(* IEC 61131-3 sources: virtual-bottling-plant/plc/src/generated/io, 9 files *)

(* ---- IO_C501.st ---- *)
(* GENERATED by plc/scripts/gen_plc_io.py from contracts/modbus/sim-io.yaml. Do not edit by hand. *)
(* Remote I/O station C501 (Modbus unit 5). *)
PROGRAM IO_C501
  VAR_EXTERNAL
    G_In : ST_SimInputs;
    G_Out : ST_SimOutputs;
  END_VAR
  VAR
    C501_Running AT %IX100.7 : BOOL;
    C501_Jam AT %IX101.0 : BOOL;
    C501_Breakdown AT %IX101.1 : BOOL;
    LSL502_CapsEmpty AT %IX101.2 : BOOL;
    C501_Run AT %QX101.2 : BOOL;
    C501_Speed AT %IW120 : UINT;
    C501_Count_HI AT %IW121 : UINT;
    C501_Count_LO AT %IW122 : UINT;
    C501_Torque AT %IW123 : UINT;
    LT502_CapHopper AT %IW124 : UINT;
    C501_Heartbeat AT %IW125 : UINT;
    C501_SpeedSP AT %QW104 : UINT;
  END_VAR
  G_In.C501_Running := C501_Running;
  G_In.C501_Jam := C501_Jam;
  G_In.C501_Breakdown := C501_Breakdown;
  G_In.LSL502_CapsEmpty := LSL502_CapsEmpty;
  C501_Run := G_Out.C501_Run;
  G_In.C501_Speed := UINT_TO_REAL(C501_Speed);
  G_In.C501_Count := UINT_TO_UDINT(C501_Count_HI) * 65536 + UINT_TO_UDINT(C501_Count_LO);
  G_In.C501_Torque := UINT_TO_REAL(C501_Torque) / 100.0;
  G_In.LT502_CapHopper := UINT_TO_REAL(LT502_CapHopper) / 10.0;
  G_In.C501_Heartbeat := C501_Heartbeat;
  C501_SpeedSP := REAL_TO_UINT(LIMIT(0.0, G_Out.C501_SpeedSP, 65535.0));
END_PROGRAM

(* ---- IO_F401.st ---- *)
(* GENERATED by plc/scripts/gen_plc_io.py from contracts/modbus/sim-io.yaml. Do not edit by hand. *)
(* Remote I/O station F401 (Modbus unit 4). *)
PROGRAM IO_F401
  VAR_EXTERNAL
    G_In : ST_SimInputs;
    G_Out : ST_SimOutputs;
  END_VAR
  VAR
    F401_Running AT %IX100.5 : BOOL;
    F401_NozzleLeak AT %IX100.6 : BOOL;
    F401_Run AT %QX101.1 : BOOL;
    F401_Speed AT %IW116 : UINT;
    F401_Count_HI AT %IW117 : UINT;
    F401_Count_LO AT %IW118 : UINT;
    F401_Heartbeat AT %IW119 : UINT;
    F401_SpeedSP AT %QW102 : UINT;
    F401_FillTargetG AT %QW103 : UINT;
  END_VAR
  G_In.F401_Running := F401_Running;
  G_In.F401_NozzleLeak := F401_NozzleLeak;
  F401_Run := G_Out.F401_Run;
  G_In.F401_Speed := UINT_TO_REAL(F401_Speed);
  G_In.F401_Count := UINT_TO_UDINT(F401_Count_HI) * 65536 + UINT_TO_UDINT(F401_Count_LO);
  G_In.F401_Heartbeat := F401_Heartbeat;
  F401_SpeedSP := REAL_TO_UINT(LIMIT(0.0, G_Out.F401_SpeedSP, 65535.0));
  F401_FillTargetG := REAL_TO_UINT(LIMIT(0.0, G_Out.F401_FillTargetG * 10.0, 65535.0));
END_PROGRAM

(* ---- IO_K801.st ---- *)
(* GENERATED by plc/scripts/gen_plc_io.py from contracts/modbus/sim-io.yaml. Do not edit by hand. *)
(* Remote I/O station K801 (Modbus unit 8). *)
PROGRAM IO_K801
  VAR_EXTERNAL
    G_In : ST_SimInputs;
    G_Out : ST_SimOutputs;
  END_VAR
  VAR
    K801_Running AT %IX102.0 : BOOL;
    K801_Jam AT %IX102.1 : BOOL;
    K801_Breakdown AT %IX102.2 : BOOL;
    K801_Run AT %QX101.5 : BOOL;
    K801_Speed AT %IW177 : UINT;
    K801_CaseCount_HI AT %IW178 : UINT;
    K801_CaseCount_LO AT %IW179 : UINT;
    K801_Heartbeat AT %IW180 : UINT;
    K801_SpeedSP AT %QW108 : UINT;
  END_VAR
  G_In.K801_Running := K801_Running;
  G_In.K801_Jam := K801_Jam;
  G_In.K801_Breakdown := K801_Breakdown;
  K801_Run := G_Out.K801_Run;
  G_In.K801_Speed := UINT_TO_REAL(K801_Speed);
  G_In.K801_CaseCount := UINT_TO_UDINT(K801_CaseCount_HI) * 65536 + UINT_TO_UDINT(K801_CaseCount_LO);
  G_In.K801_Heartbeat := K801_Heartbeat;
  K801_SpeedSP := REAL_TO_UINT(LIMIT(0.0, G_Out.K801_SpeedSP, 65535.0));
END_PROGRAM

(* ---- IO_L601.st ---- *)
(* GENERATED by plc/scripts/gen_plc_io.py from contracts/modbus/sim-io.yaml. Do not edit by hand. *)
(* Remote I/O station L601 (Modbus unit 6). *)
PROGRAM IO_L601
  VAR_EXTERNAL
    G_In : ST_SimInputs;
    G_Out : ST_SimOutputs;
  END_VAR
  VAR
    L601_Running AT %IX101.3 : BOOL;
    L601_RollEmpty AT %IX101.4 : BOOL;
    L601_LabelError AT %IX101.5 : BOOL;
    L601_Breakdown AT %IX101.6 : BOOL;
    L601_Run AT %QX101.3 : BOOL;
    L601_Speed AT %IW126 : UINT;
    L601_Count_HI AT %IW127 : UINT;
    L601_Count_LO AT %IW128 : UINT;
    L601_RollRemaining AT %IW129 : UINT;
    L601_Heartbeat AT %IW130 : UINT;
    L601_SpeedSP AT %QW105 : UINT;
  END_VAR
  G_In.L601_Running := L601_Running;
  G_In.L601_RollEmpty := L601_RollEmpty;
  G_In.L601_LabelError := L601_LabelError;
  G_In.L601_Breakdown := L601_Breakdown;
  L601_Run := G_Out.L601_Run;
  G_In.L601_Speed := UINT_TO_REAL(L601_Speed);
  G_In.L601_Count := UINT_TO_UDINT(L601_Count_HI) * 65536 + UINT_TO_UDINT(L601_Count_LO);
  G_In.L601_RollRemaining := UINT_TO_REAL(L601_RollRemaining);
  G_In.L601_Heartbeat := L601_Heartbeat;
  L601_SpeedSP := REAL_TO_UINT(LIMIT(0.0, G_Out.L601_SpeedSP, 65535.0));
END_PROGRAM

(* ---- IO_LINE.st ---- *)
(* GENERATED by plc/scripts/gen_plc_io.py from contracts/modbus/sim-io.yaml. Do not edit by hand. *)
(* Remote I/O station LINE (Modbus unit 9). *)
PROGRAM IO_LINE
  VAR_EXTERNAL
    G_In : ST_SimInputs;
  END_VAR
  VAR
    CV1_Full AT %IX102.3 : BOOL;
    CV2_Full AT %IX102.4 : BOOL;
    CV3_Full AT %IX102.5 : BOOL;
    CV4_Full AT %IX102.6 : BOOL;
    PB_Start AT %IX102.7 : BOOL;
    PB_Stop AT %IX103.0 : BOOL;
    PB_Reset AT %IX103.1 : BOOL;
    SIM_TimeMs_HI AT %IW181 : UINT;
    SIM_TimeMs_LO AT %IW182 : UINT;
    CV1_Fill AT %IW183 : UINT;
    CV2_Fill AT %IW184 : UINT;
    CV3_Fill AT %IW185 : UINT;
    CV4_Fill AT %IW186 : UINT;
    LINE_Heartbeat AT %IW187 : UINT;
  END_VAR
  G_In.CV1_Full := CV1_Full;
  G_In.CV2_Full := CV2_Full;
  G_In.CV3_Full := CV3_Full;
  G_In.CV4_Full := CV4_Full;
  G_In.PB_Start := PB_Start;
  G_In.PB_Stop := PB_Stop;
  G_In.PB_Reset := PB_Reset;
  G_In.SIM_TimeMs := UINT_TO_UDINT(SIM_TimeMs_HI) * 65536 + UINT_TO_UDINT(SIM_TimeMs_LO);
  G_In.CV1_Fill := UINT_TO_REAL(CV1_Fill);
  G_In.CV2_Fill := UINT_TO_REAL(CV2_Fill);
  G_In.CV3_Fill := UINT_TO_REAL(CV3_Fill);
  G_In.CV4_Fill := UINT_TO_REAL(CV4_Fill);
  G_In.LINE_Heartbeat := LINE_Heartbeat;
END_PROGRAM

(* ---- IO_P201.st ---- *)
(* GENERATED by plc/scripts/gen_plc_io.py from contracts/modbus/sim-io.yaml. Do not edit by hand. *)
(* Remote I/O station P201 (Modbus unit 2). *)
PROGRAM IO_P201
  VAR_EXTERNAL
    G_In : ST_SimInputs;
    G_Out : ST_SimOutputs;
  END_VAR
  VAR
    ZS203_DivertOpen AT %IX100.3 : BOOL;
    XV203_Divert AT %QX100.7 : BOOL;
    TT201_InTemp AT %IW109 : UINT;
    TT202_OutTemp AT %IW110 : UINT;
    FT201_Flow AT %IW111 : UINT;
    PT201_SteamPressure AT %IW112 : UINT;
    P201_Heartbeat AT %IW113 : UINT;
    TCV201_SteamValve AT %QW101 : UINT;
  END_VAR
  G_In.ZS203_DivertOpen := ZS203_DivertOpen;
  XV203_Divert := G_Out.XV203_Divert;
  G_In.TT201_InTemp := UINT_TO_REAL(TT201_InTemp) / 10.0;
  G_In.TT202_OutTemp := UINT_TO_REAL(TT202_OutTemp) / 10.0;
  G_In.FT201_Flow := UINT_TO_REAL(FT201_Flow);
  G_In.PT201_SteamPressure := UINT_TO_REAL(PT201_SteamPressure) / 100.0;
  G_In.P201_Heartbeat := P201_Heartbeat;
  TCV201_SteamValve := REAL_TO_UINT(LIMIT(0.0, G_Out.TCV201_SteamValve * 10.0, 65535.0));
END_PROGRAM

(* ---- IO_Q701.st ---- *)
(* GENERATED by plc/scripts/gen_plc_io.py from contracts/modbus/sim-io.yaml. Do not edit by hand. *)
(* Remote I/O station Q701 (Modbus unit 7). *)
PROGRAM IO_Q701
  VAR_EXTERNAL
    G_In : ST_SimInputs;
    G_Out : ST_SimOutputs;
  END_VAR
  VAR
    Q701_Running AT %IX101.7 : BOOL;
    Q701_Run AT %QX101.4 : BOOL;
    Q701_Speed AT %IW131 : UINT;
    Q701_Count_HI AT %IW132 : UINT;
    Q701_Count_LO AT %IW133 : UINT;
    Q701_RejectCount_HI AT %IW134 : UINT;
    Q701_RejectCount_LO AT %IW135 : UINT;
    WT701_LastWeight AT %IW136 : UINT;
    Q701_Heartbeat AT %IW137 : UINT;
    Q701_N01_Seq AT %IW141 : UINT;
    Q701_N01_Mean AT %IW142 : UINT;
    Q701_N01_Range AT %IW143 : UINT;
    Q701_N02_Seq AT %IW144 : UINT;
    Q701_N02_Mean AT %IW145 : UINT;
    Q701_N02_Range AT %IW146 : UINT;
    Q701_N03_Seq AT %IW147 : UINT;
    Q701_N03_Mean AT %IW148 : UINT;
    Q701_N03_Range AT %IW149 : UINT;
    Q701_N04_Seq AT %IW150 : UINT;
    Q701_N04_Mean AT %IW151 : UINT;
    Q701_N04_Range AT %IW152 : UINT;
    Q701_N05_Seq AT %IW153 : UINT;
    Q701_N05_Mean AT %IW154 : UINT;
    Q701_N05_Range AT %IW155 : UINT;
    Q701_N06_Seq AT %IW156 : UINT;
    Q701_N06_Mean AT %IW157 : UINT;
    Q701_N06_Range AT %IW158 : UINT;
    Q701_N07_Seq AT %IW159 : UINT;
    Q701_N07_Mean AT %IW160 : UINT;
    Q701_N07_Range AT %IW161 : UINT;
    Q701_N08_Seq AT %IW162 : UINT;
    Q701_N08_Mean AT %IW163 : UINT;
    Q701_N08_Range AT %IW164 : UINT;
    Q701_N09_Seq AT %IW165 : UINT;
    Q701_N09_Mean AT %IW166 : UINT;
    Q701_N09_Range AT %IW167 : UINT;
    Q701_N10_Seq AT %IW168 : UINT;
    Q701_N10_Mean AT %IW169 : UINT;
    Q701_N10_Range AT %IW170 : UINT;
    Q701_N11_Seq AT %IW171 : UINT;
    Q701_N11_Mean AT %IW172 : UINT;
    Q701_N11_Range AT %IW173 : UINT;
    Q701_N12_Seq AT %IW174 : UINT;
    Q701_N12_Mean AT %IW175 : UINT;
    Q701_N12_Range AT %IW176 : UINT;
    Q701_SpeedSP AT %QW106 : UINT;
    Q701_RejectLimitG AT %QW107 : UINT;
  END_VAR
  G_In.Q701_Running := Q701_Running;
  Q701_Run := G_Out.Q701_Run;
  G_In.Q701_Speed := UINT_TO_REAL(Q701_Speed);
  G_In.Q701_Count := UINT_TO_UDINT(Q701_Count_HI) * 65536 + UINT_TO_UDINT(Q701_Count_LO);
  G_In.Q701_RejectCount := UINT_TO_UDINT(Q701_RejectCount_HI) * 65536 + UINT_TO_UDINT(Q701_RejectCount_LO);
  G_In.WT701_LastWeight := UINT_TO_REAL(WT701_LastWeight) / 10.0;
  G_In.Q701_Heartbeat := Q701_Heartbeat;
  G_In.Q701_N01_Seq := Q701_N01_Seq;
  G_In.Q701_N01_Mean := UINT_TO_REAL(Q701_N01_Mean) / 10.0;
  G_In.Q701_N01_Range := UINT_TO_REAL(Q701_N01_Range) / 10.0;
  G_In.Q701_N02_Seq := Q701_N02_Seq;
  G_In.Q701_N02_Mean := UINT_TO_REAL(Q701_N02_Mean) / 10.0;
  G_In.Q701_N02_Range := UINT_TO_REAL(Q701_N02_Range) / 10.0;
  G_In.Q701_N03_Seq := Q701_N03_Seq;
  G_In.Q701_N03_Mean := UINT_TO_REAL(Q701_N03_Mean) / 10.0;
  G_In.Q701_N03_Range := UINT_TO_REAL(Q701_N03_Range) / 10.0;
  G_In.Q701_N04_Seq := Q701_N04_Seq;
  G_In.Q701_N04_Mean := UINT_TO_REAL(Q701_N04_Mean) / 10.0;
  G_In.Q701_N04_Range := UINT_TO_REAL(Q701_N04_Range) / 10.0;
  G_In.Q701_N05_Seq := Q701_N05_Seq;
  G_In.Q701_N05_Mean := UINT_TO_REAL(Q701_N05_Mean) / 10.0;
  G_In.Q701_N05_Range := UINT_TO_REAL(Q701_N05_Range) / 10.0;
  G_In.Q701_N06_Seq := Q701_N06_Seq;
  G_In.Q701_N06_Mean := UINT_TO_REAL(Q701_N06_Mean) / 10.0;
  G_In.Q701_N06_Range := UINT_TO_REAL(Q701_N06_Range) / 10.0;
  G_In.Q701_N07_Seq := Q701_N07_Seq;
  G_In.Q701_N07_Mean := UINT_TO_REAL(Q701_N07_Mean) / 10.0;
  G_In.Q701_N07_Range := UINT_TO_REAL(Q701_N07_Range) / 10.0;
  G_In.Q701_N08_Seq := Q701_N08_Seq;
  G_In.Q701_N08_Mean := UINT_TO_REAL(Q701_N08_Mean) / 10.0;
  G_In.Q701_N08_Range := UINT_TO_REAL(Q701_N08_Range) / 10.0;
  G_In.Q701_N09_Seq := Q701_N09_Seq;
  G_In.Q701_N09_Mean := UINT_TO_REAL(Q701_N09_Mean) / 10.0;
  G_In.Q701_N09_Range := UINT_TO_REAL(Q701_N09_Range) / 10.0;
  G_In.Q701_N10_Seq := Q701_N10_Seq;
  G_In.Q701_N10_Mean := UINT_TO_REAL(Q701_N10_Mean) / 10.0;
  G_In.Q701_N10_Range := UINT_TO_REAL(Q701_N10_Range) / 10.0;
  G_In.Q701_N11_Seq := Q701_N11_Seq;
  G_In.Q701_N11_Mean := UINT_TO_REAL(Q701_N11_Mean) / 10.0;
  G_In.Q701_N11_Range := UINT_TO_REAL(Q701_N11_Range) / 10.0;
  G_In.Q701_N12_Seq := Q701_N12_Seq;
  G_In.Q701_N12_Mean := UINT_TO_REAL(Q701_N12_Mean) / 10.0;
  G_In.Q701_N12_Range := UINT_TO_REAL(Q701_N12_Range) / 10.0;
  Q701_SpeedSP := REAL_TO_UINT(LIMIT(0.0, G_Out.Q701_SpeedSP, 65535.0));
  Q701_RejectLimitG := REAL_TO_UINT(LIMIT(0.0, G_Out.Q701_RejectLimitG * 10.0, 65535.0));
END_PROGRAM

(* ---- IO_T101.st ---- *)
(* GENERATED by plc/scripts/gen_plc_io.py from contracts/modbus/sim-io.yaml. Do not edit by hand. *)
(* Remote I/O station T101 (Modbus unit 1). *)
PROGRAM IO_T101
  VAR_EXTERNAL
    G_In : ST_SimInputs;
    G_Out : ST_SimOutputs;
  END_VAR
  VAR
    LSL101_Empty AT %IX100.0 : BOOL;
    M101_Running AT %IX100.1 : BOOL;
    T101_CipDone AT %IX100.2 : BOOL;
    XV101_Water AT %QX100.0 : BOOL;
    XV102_Conc AT %QX100.1 : BOOL;
    XV103_Sugar AT %QX100.2 : BOOL;
    M101_Agitator AT %QX100.3 : BOOL;
    P101_TransferPump AT %QX100.4 : BOOL;
    XV109_Drain AT %QX100.5 : BOOL;
    T101_CipRun AT %QX100.6 : BOOL;
    LT101_Level AT %IW100 : UINT;
    AT101_Brix AT %IW101 : UINT;
    FT101_WaterFlow AT %IW102 : UINT;
    FT102_ConcFlow AT %IW103 : UINT;
    FT103_SugarFlow AT %IW104 : UINT;
    ST101_AgitatorRpm AT %IW105 : UINT;
    T101_ConcLotNo_HI AT %IW106 : UINT;
    T101_ConcLotNo_LO AT %IW107 : UINT;
    T101_Heartbeat AT %IW108 : UINT;
    T101_ConcSelect AT %QW100 : UINT;
  END_VAR
  G_In.LSL101_Empty := LSL101_Empty;
  G_In.M101_Running := M101_Running;
  G_In.T101_CipDone := T101_CipDone;
  XV101_Water := G_Out.XV101_Water;
  XV102_Conc := G_Out.XV102_Conc;
  XV103_Sugar := G_Out.XV103_Sugar;
  M101_Agitator := G_Out.M101_Agitator;
  P101_TransferPump := G_Out.P101_TransferPump;
  XV109_Drain := G_Out.XV109_Drain;
  T101_CipRun := G_Out.T101_CipRun;
  G_In.LT101_Level := UINT_TO_REAL(LT101_Level) / 10.0;
  G_In.AT101_Brix := UINT_TO_REAL(AT101_Brix) / 100.0;
  G_In.FT101_WaterFlow := UINT_TO_REAL(FT101_WaterFlow);
  G_In.FT102_ConcFlow := UINT_TO_REAL(FT102_ConcFlow);
  G_In.FT103_SugarFlow := UINT_TO_REAL(FT103_SugarFlow);
  G_In.ST101_AgitatorRpm := UINT_TO_REAL(ST101_AgitatorRpm);
  G_In.T101_ConcLotNo := UINT_TO_UDINT(T101_ConcLotNo_HI) * 65536 + UINT_TO_UDINT(T101_ConcLotNo_LO);
  G_In.T101_Heartbeat := T101_Heartbeat;
  T101_ConcSelect := REAL_TO_UINT(LIMIT(0.0, G_Out.T101_ConcSelect, 65535.0));
END_PROGRAM

(* ---- IO_T301.st ---- *)
(* GENERATED by plc/scripts/gen_plc_io.py from contracts/modbus/sim-io.yaml. Do not edit by hand. *)
(* Remote I/O station T301 (Modbus unit 3). *)
PROGRAM IO_T301
  VAR_EXTERNAL
    G_In : ST_SimInputs;
    G_Out : ST_SimOutputs;
  END_VAR
  VAR
    LSL301_Low AT %IX100.4 : BOOL;
    XV309_Drain AT %QX101.0 : BOOL;
    LT301_Level AT %IW114 : UINT;
    T301_Heartbeat AT %IW115 : UINT;
  END_VAR
  G_In.LSL301_Low := LSL301_Low;
  XV309_Drain := G_Out.XV309_Drain;
  G_In.LT301_Level := UINT_TO_REAL(LT301_Level) / 10.0;
  G_In.T301_Heartbeat := T301_Heartbeat;
END_PROGRAM
